Fanuc KAREL source: KA00220.KL

PROGRAM KA00220
%NOLOCKGROUP
VAR
  SRC: ARRAY[4] OF JOINTPOS
  DST: ARRAY[4] OF STRING[20]
BEGIN
  DST = SRC
END KA00220
